(* IEC 61131-3 sources: daoli-st-library/DL_MathData (part 17) *)

(* ---- FC_DL_LinearScale.st ---- *)
(*==============================================================================
 * 组件名称 (Component)  : FC_DL_LinearScale
 * 所属子库 (Sublibrary) : DL_MathData
 * 当前版本 (Version)    : 1.0.0
 * 兼容性   (Platform)   : CODESYS 3.5 / TwinCAT 3 / 汇川 InoProShop / Machine Expert
 *                         仅依赖 Standard.library（ABS / MIN / MAX），全 REAL 运算
 * 功能描述 (Function)   : 模拟量原始码 → 工程量的线性标定。如 0..27648 对应 0..1.6MPa，
 *                         或 4..20mA 对应 0..100%。内置量程为零防御（除零保护）、
 *                         反向量程支持、输出双侧钳位、输入占量程百分比输出。
 *                         钳位判定使用浮点容差，不做浮点判等。
 * 开源溯源 (Origin)     : 原创实现。防御结构与模板库 05-algorithm-templates.md
 *                         的 FC_LinearScale 思路同源，按本库故障码体系重写并加严。
 * 依赖     (Depends)    : 无 DL_ 内部依赖
 * 说明     (Note)       : NaN / Inf 检测在纯 IEC 61131-3 中无标准手段（各平台对
 *                         比较运算返回值处理不一致），故 v1.0.0 不做该检测，
 *                         故障码 16#0001_0006 预留给支持 NaN 检测的平台版本。
 * 红线自检 (Redline)    : R1 ✓ 零全局变量表与外部变量引用 ｜ R2 ✓ 零物理 IO 地址直写
 *                         R3 ✓ 纯 IEC 61131-3 ｜ R4 ✓ 除零/排序/双侧钳位/容差判等（本轮 R4 样板）
 *                         R5 ✓ 全变量中英双语同行注释 ｜ R6 N/A（无状态机）｜ R7 N/A（无实例调用）
 * 修订历史 (Revision)   :
 *   2026-11-14  v1.0.0  首版入库（Phase 1 冷启动 · Level 0 批次）
 *============================================================================*)
FUNCTION FC_DL_LinearScale : REAL
VAR_INPUT
    fIn      : REAL;                 // 原始输入值 [raw] / Raw input value [raw]
    fInMin   : REAL := 0.0;          // 输入量程下限 [raw] / Input range low [raw]
    fInMax   : REAL := 27648.0;      // 输入量程上限 [raw] / Input range high [raw]
    fOutMin  : REAL := 0.0;          // 工程量下限 [EU] / Engineering range low [EU]
    fOutMax  : REAL := 100.0;        // 工程量上限 [EU] / Engineering range high [EU]
    bClamp   : BOOL := TRUE;         // 是否双侧钳位到工程量程 / Enable two-sided clamping
END_VAR
VAR_OUTPUT
    bValid   : BOOL;                 // 换算有效标志，FALSE 表示量程非法 / Conversion valid flag, FALSE means invalid range
    bClamped : BOOL;                 // 结果被钳位标志 / Result clamped flag
    fPercent : REAL;                 // 输入占量程百分比 [%]，可超 0..100 / Input as percent of span [%], may exceed 0..100
    uErrorId : UDINT;                // 故障码，0 = 无故障 / Error code, 0 = no error
END_VAR
VAR
    fSpanIn  : REAL;                 // 输入量程跨度 [raw]，可为负（反向标定） / Input span [raw], negative for reverse scaling
    fSpanOut : REAL;                 // 输出量程跨度 [EU]，可为负 / Output span [EU], may be negative
    fResult  : REAL;                 // 中间结果 [EU] / Intermediate result [EU]
    fNorm    : REAL;                 // 归一化比值 [0..1 附近]，无量纲 / Normalized ratio, dimensionless
    fOutLo   : REAL;                 // 输出下限，已排序 [EU] / Ordered output low limit [EU]
    fOutHi   : REAL;                 // 输出上限，已排序 [EU] / Ordered output high limit [EU]
    fBefore  : REAL;                 // 钳位前的结果快照，用于判定是否发生钳位 [EU] / Pre-clamp snapshot [EU]
END_VAR
VAR CONSTANT
    DL_FLOAT_EPS : REAL := 1.0E-6;   // 浮点判零容差 / Float zero tolerance
END_VAR

(*------------------------------------------------------------------------------
 * 段 1｜安全预置：任何异常路径下返回值落到工程量下限
 *      Safe preset: on every error path the return value falls back to the output low
 *-----------------------------------------------------------------------------*)
FC_DL_LinearScale := fOutMin;
bValid            := TRUE;
bClamped          := FALSE;
fPercent          := 0.0;
uErrorId          := 16#0000_0000;
fResult           := fOutMin;
fBefore           := fOutMin;

(*------------------------------------------------------------------------------
 * 段 2｜量程跨度计算 + 防除零（边界 B1 / B6）
 *      Span computation and divide-by-zero guard
 *      浮点判零用 ABS(..) <= EPS，禁止 fSpanIn = 0.0
 *      该段必须先于任何除法，fPercent 的计算建立在跨度已校验的前提上
 *-----------------------------------------------------------------------------*)
fSpanIn  := fInMax - fInMin;
fSpanOut := fOutMax - fOutMin;

IF ABS(fSpanIn) <= DL_FLOAT_EPS THEN
    bValid            := FALSE;
    uErrorId          := 16#0001_0002;
    FC_DL_LinearScale := fOutMin;
    RETURN;
END_IF

(*------------------------------------------------------------------------------
 * 段 3｜归一化与百分比（边界 B2）：反向量程天然支持
 *      Normalization and percentage: reverse ranges are supported by construction
 *      fInMax < fInMin 时 fSpanIn 为负，比值自动反向，0% 落在 fInMax 侧
 *-----------------------------------------------------------------------------*)
fNorm    := (fIn - fInMin) / fSpanIn;
fPercent := fNorm * 100.0;
fResult  := fOutMin + fNorm * fSpanOut;

(*------------------------------------------------------------------------------
 * 段 4｜输出边界排序（边界 B3）：钳位前必须先排序
 *      Output limit ordering before clamping
 *      若输出量程传反而不排序，钳位会把结果压到错误端点，现象是"钳位看似
 *      生效而输出全错"，这是本组件最隐蔽的失效模式
 *-----------------------------------------------------------------------------*)
fOutLo := MIN(fOutMin, fOutMax);
fOutHi := MAX(fOutMin, fOutMax);

(*------------------------------------------------------------------------------
 * 段 5｜双侧钳位（边界 B4/B5）：上下限成对出现，只用一侧是安全红线错误
 *      Two-sided clamping: both limits are mandatory, one-sided is a safety defect
 *      只做上限会让负向冲击直接打穿执行机构；钳位判定用容差而非不等号
 *-----------------------------------------------------------------------------*)
IF bClamp THEN
    fBefore := fResult;

    IF fResult < fOutLo THEN
        fResult := fOutLo;
    ELSIF fResult > fOutHi THEN
        fResult := fOutHi;
    END_IF

    IF ABS(fResult - fBefore) > DL_FLOAT_EPS THEN
        bClamped := TRUE;
    END_IF
END_IF

(*------------------------------------------------------------------------------
 * 段 6｜结果回写（边界 B7）：字面量均带小数点，全程 REAL，不混入 LREAL
 *      Result write-back: literals carry decimal points, REAL stays REAL
 *-----------------------------------------------------------------------------*)
FC_DL_LinearScale := fResult;
END_FUNCTION

(* ---- FC_DL_LineIntersection.st ---- *)
(*==============================================================================
 * 组件名称 (Component)  : FC_DL_LineIntersection
 * 所属子库 (Sublibrary) : DL_MathData
 * 当前版本 (Version)    : 1.0.0
 * 兼容性   (Platform)   : CODESYS 3.5 / TwinCAT 3 / 汇川 InoProShop / Machine Expert
 *                         仅依赖 Standard.library（ABS），全 LREAL 运算，无状态
 * 功能描述 (Function)   : 二维两直线（或两线段）交点求解。返回"是否存在唯一交点"的布尔量，
 *                         交点坐标与两个线段参数经状态输出给出，双通道并存的目的是让调用方
 *                         既能直接用作条件判断，也能拿到参数做端点命中判据。
 *                         用于视觉十字标定、皮带跑偏中心线求交、两台相机视场交叠区定位、
 *                         机器人平面两轴交汇点计算。
 *
 * 【失真与语义披露 / Distortion disclosure】
 *   1) 线段模式返回 FALSE 时 uErrorId = 0：业务上的"两段不相交"是正常判定结果，
 *      不是故障。若也置故障码，上位机会把正常判定当异常刷屏，真正的配置错误就被淹了。
 *   2) 重合直线归入平行类（16#0002_000D）：无穷多交点无法用单一坐标表达，
 *      与其随机给一个点，不如明确说"没有唯一交点"。线段模式下"平行且不共线"的两段
 *      永远不可能相交，属于正常业务判定，返回 FALSE 且不置码；只有重合（共线）才报码。
 *   3) 平行判据用绝对容差，而坐标量级到 1e6 时行列式 fDen 可到 1e12，因此 fEps 必须
 *      按坐标量级配置，经验式 fEps ≈ 1e-9 × 坐标量级²。用 1e-9 去判 1e12 量级的行列式，
 *      等于把平行判据关掉了。
 *   4) 本函数不检测 NaN/Inf：IEC 61131-3 无标准判据，强行判断会引入编译器方言。
 *
 * 开源溯源 (Origin)     : 原创实现（参考西门子 LGF 数学功能组中平面几何族的分类位置，
 *                         解析几何求交为公开数学方法，clean-room 独立实现）
 * 依赖     (Depends)    : 无 DL_ 内部依赖；Standard.library: ABS
 * 红线自检 (Redline)    : R1 ✓ 零全局变量表与外部变量引用 ｜ R2 ✓ 零物理 IO 地址直写
 *                         R3 ✓ 纯 IEC 61131-3（无指针、无厂商私有符号）
 *                         R4 ✓ 零长度线判据 + 容差规整 + 行列式判零 + 无交点显式清 0
 *                         R5 ✓ 全变量中英双语同行注释 ｜ R6 N/A（无状态机）｜ R7 N/A（无实例调用）
 * 修订历史 (Revision)   :
 *   2026-11-14  v1.0.0  首版入库（Phase 1 收口批次 · R3）
 *============================================================================*)
FUNCTION FC_DL_LineIntersection : BOOL
VAR_INPUT
    fX1         : LREAL;                  // 线 1 起点 X [mm] / Line 1 start X [mm]
    fY1         : LREAL;                  // 线 1 起点 Y [mm] / Line 1 start Y [mm]
    fX2         : LREAL;                  // 线 1 终点 X [mm] / Line 1 end X [mm]
    fY2         : LREAL;                  // 线 1 终点 Y [mm] / Line 1 end Y [mm]
    fX3         : LREAL;                  // 线 2 起点 X [mm] / Line 2 start X [mm]
    fY3         : LREAL;                  // 线 2 起点 Y [mm] / Line 2 start Y [mm]
    fX4         : LREAL;                  // 线 2 终点 X [mm] / Line 2 end X [mm]
    fY4         : LREAL;                  // 线 2 终点 Y [mm] / Line 2 end Y [mm]
    fEps        : LREAL := 1.0E-9;        // 平行判定容差（须按坐标量级配置）/ Parallel tolerance, scale with the coordinate range
    bSegmentMode: BOOL := FALSE;          // TRUE = 按线段求交，交点须落在两段内 / TRUE = segment mode
END_VAR
VAR_OUTPUT
    fX       : LREAL;                     // 交点 X [mm]，无交点时为 0 / Intersection X [mm], 0 when none
    fY       : LREAL;                     // 交点 Y [mm]，无交点时为 0 / Intersection Y [mm], 0 when none
    fT       : LREAL;                     // 线 1 参数 t，0 = 起点、1 = 终点 / Parameter along line 1
    fU       : LREAL;                     // 线 2 参数 u，0 = 起点、1 = 终点 / Parameter along line 2
    uErrorId : UDINT;                     // 故障码，0 = 无故障 / Error code, 0 = no error
END_VAR
VAR
    fDen  : LREAL;                        // 行列式分母 / Determinant denominator
    fDx1  : LREAL;                        // 线 1 方向 X 分量 [mm] / Line 1 direction X [mm]
    fDy1  : LREAL;                        // 线 1 方向 Y 分量 [mm] / Line 1 direction Y [mm]
    fDx2  : LREAL;                        // 线 2 方向 X 分量 [mm] / Line 2 direction X [mm]
    fDy2  : LREAL;                        // 线 2 方向 Y 分量 [mm] / Line 2 direction Y [mm]
    fEpsEff : LREAL;                      // 规整后的容差 / Normalised tolerance
    fTol  : LREAL;                        // 线段模式的参数区间容差 / Parameter tolerance in segment mode
    fNumT : LREAL;                        // t 的分子 / Numerator of t
    fNumU : LREAL;                        // u 的分子 / Numerator of u
    bLineDegenerate : BOOL;               // 任一线退化为点（起终点重合）/ Either line degenerated to a point
    bCoincident : BOOL;                   // 两线共线（重合），平行判定后的细分 / The two lines are coincident
END_VAR
VAR CONSTANT
    DL_LI_DEADBAND : LREAL := 1.0E-6;     // 零长度线判定容差 [mm] / Zero-length line tolerance [mm]
    DL_LI_EPS_MIN  : LREAL := 1.0E-12;    // 容差下限，防止把容差填成 0 / Tolerance floor
END_VAR

(*------------------------------------------------------------------------------
 * 段 1｜安全预置（边界 B6）：无交点时输出必须显式清 0，禁止依赖"局部变量默认值"
 *      Safe preset: outputs are explicitly zeroed, local defaults are never trusted
 *      部分平台的 FC 局部变量不保证每拍复位，靠默认值会让上一次的交点粘住
 *-----------------------------------------------------------------------------*)
FC_DL_LineIntersection := FALSE;
fX       := 0.0;
fY       := 0.0;
fT       := 0.0;
fU       := 0.0;
uErrorId := 16#0000_0000;

(*------------------------------------------------------------------------------
 * 段 2｜退化线检测（边界 B2）：起点终点重合/填反是最常见的标定配置错误，必须报码
 *      Degenerate-line check: start equal to end is the most common calibration mistake
 *      用曼哈顿距离判零长度：比平方和开方便宜，且对 LREAL 无溢出风险
 *-----------------------------------------------------------------------------*)
bLineDegenerate := ((ABS(fX2 - fX1) + ABS(fY2 - fY1)) <= DL_LI_DEADBAND)
                   OR ((ABS(fX4 - fX3) + ABS(fY4 - fY3)) <= DL_LI_DEADBAND);

IF bLineDegenerate THEN
    uErrorId := 16#0001_0001;
    RETURN;
END_IF

(*------------------------------------------------------------------------------
 * 段 3｜容差规整（边界 B1）：容差不能为 0 或负，否则平行判据失效
 *      Tolerance normalisation: zero or negative would disable the parallel test
 *-----------------------------------------------------------------------------*)
fEpsEff := fEps;

IF fEpsEff <= 0.0 THEN
    fEpsEff  := 1.0E-9;
    uErrorId := 16#0001_0001;
END_IF

IF fEpsEff < DL_LI_EPS_MIN THEN
    fEpsEff := DL_LI_EPS_MIN;
END_IF

(*------------------------------------------------------------------------------
 * 段 4｜方向向量与行列式（边界 B5）：分母只算一次，两条参数方程共用
 *      Direction vectors and determinant, computed once for both parametric equations
 *-----------------------------------------------------------------------------*)
fDx1 := fX2 - fX1;
fDy1 := fY2 - fY1;
fDx2 := fX4 - fX3;
fDy2 := fY4 - fY3;

fDen := (fDx1 * fDy2) - (fDy1 * fDx2);

(*------------------------------------------------------------------------------
 * 段 5｜平行/重合判定（边界 B3/B4）：无唯一交点
 *      Parallel or coincident: no unique intersection
 *      线段模式下"平行且不共线"的两段永远不相交，属正常业务判定，不置故障码；
 *      重合则有无穷多交点，仍是配置/数据问题，必须报码
 *      In segment mode, parallel non-collinear segments are a normal verdict, not a fault
 *-----------------------------------------------------------------------------*)
IF ABS(fDen) <= fEpsEff THEN

    bCoincident := (ABS(((fX3 - fX1) * fDy1) - ((fY3 - fY1) * fDx1)) <= fEpsEff);

    IF bSegmentMode AND (NOT bCoincident) THEN
        RETURN;
    END_IF

    uErrorId := 16#0002_000D;
    RETURN;

END_IF

(*------------------------------------------------------------------------------
 * 段 6｜参数求解：克拉默法则，分母在段 5 已判非零
 *      Parameter solution by Cramer's rule, the denominator was proven non-zero
 *-----------------------------------------------------------------------------*)
fNumT := (((fX3 - fX1) * fDy2) - ((fY3 - fY1) * fDx2));
fNumU := (((fX3 - fX1) * fDy1) - ((fY3 - fY1) * fDx1));

fT := fNumT / fDen;
fU := fNumU / fDen;

(*------------------------------------------------------------------------------
 * 段 7｜线段模式判定（边界 B3）：交点须落在两段的参数区间内
 *      Segment mode: the intersection must lie inside both parameter ranges
 *      端点命中算相交（容差取 fEpsEff 量级），否则相邻两段共端点时会被判成"不相交"；
 *      判定失败时 fT / fU 保留实际参数，便于上位机判断"差多远"，但坐标清 0
 *-----------------------------------------------------------------------------*)
IF bSegmentMode THEN

    fTol := fEpsEff;

    IF (fT < (0.0 - fTol)) OR (fT > (1.0 + fTol)) THEN
        (* 业务判定，不置故障码：线段不相交是正常结果 *)
        (* A business verdict, not a fault: disjoint segments are perfectly normal *)
        RETURN;
    END_IF

    IF (fU < (0.0 - fTol)) OR (fU > (1.0 + fTol)) THEN
        RETURN;
    END_IF

END_IF

(*------------------------------------------------------------------------------
 * 段 8｜交点求值（边界 B5）：一律由线 1 参数化，两式取平均会多引入一次误差
 *      Evaluate with line 1 only: averaging both equations adds error instead of removing it
 *-----------------------------------------------------------------------------*)
fX := fX1 + (fT * fDx1);
fY := fY1 + (fT * fDy1);

FC_DL_LineIntersection := TRUE;
END_FUNCTION

(* ---- FC_DL_LintToDintSat.st ---- *)
(*
    FC_DL_LintToDintSat —— LINT 到 DINT 双向域外饱和转换
    ------------------------------------------------------------------
    分类      : DL_MathData / Convert
    前缀      : FC_DL_
    版本      : 1.0.0
    溯源      : IEC 61131-3 标准语义的道莅防御性实现
                （接口语义由 IEC 61131-3 定义，内部委托平台内建 LINT_TO_DINT，
                  外围统一错误码 / 钳位 / 双语文档；clean-room 重写，
                  未复制任何闭源厂商源码，参考实现仅限 MIT/Apache 许可）
    平台      : 纯 IEC 61131-3，CODESYS / TwinCAT / InoProShop 通用
    作者      : 道莅代码库 · PLC编程专家（R17）
    ------------------------------------------------------------------
    功能说明  : 将 LINT 防御性转换为 DINT 并作为返回值输出，域内转换委托平台内建 LINT_TO_DINT；
                nIn 超 DINT 上界 2147483647 时饱和输出 2147483647 并置信息级 16#0001_0200；
                nIn 低于 DINT 下界 −2147483648 时饱和输出 −2147483648 并置信息级 16#0001_022D；
                下界输出采用计算式 -DL_DINT_MAX - 1，禁用负数字面量直写
                （部分编译器把负号解析为对一个越界正字面量取负，产生告警或错误结果）；
                极值比较采用双侧比较，禁用 ABS(nIn)（R55：有符号极值取绝对值会回绕漏判）；
                钳位方向：双侧饱和（−2147483648 ~ 2147483647），绝不回绕；
                纯整数域无 NaN/±INF 态，故无故障级路径（三个故障槽预留）。
    错误码    : 16#0001_0200 nIn 超 DINT 上界，已饱和至 2147483647——信息级，正常防御
                16#0001_022D nIn 低于 DINT 下界，已饱和至 −2147483648——信息级，正常防御
                16#0001_02EE 预留禁用（故障级，不得挪用）
                16#0001_02EF 预留禁用（故障级，不得挪用）
                16#0001_02F0 预留禁用（故障级，不得挪用）
    状态机    : R6 标注 N/A —— 本组件为纯函数无顺序状态机，无 CASE 可写，非法状态不可能出现，故以本节说明替代 ELSE 兜底
    修订记录  : 2026-11-16 v1.0.0 首次入库（R17）
*)
FUNCTION FC_DL_LintToDintSat : DINT
VAR_INPUT
    nIn : LINT; // 待转换 64 位有符号整数，建议域 ±9223372036854775807 [无量纲] / signed 64-bit integer to convert, suggested domain +/-9223372036854775807 [dimensionless]
END_VAR
VAR_OUTPUT
    eErr   : UDINT; // 错误码，0=正常 / error id, 0=ok
    bError : BOOL;  // 是否出错，eErr 非 0 时为 TRUE / error flag, TRUE when eErr is nonzero
    bValid : BOOL;  // 输出是否有效可用 / output valid flag
END_VAR
VAR CONSTANT
    DL_DINT_MAX_L : LINT := 2147483647;      // DINT 上界，用 LINT 承载以便域外比较 [无量纲] / DINT upper bound carried in LINT for out-of-domain comparison [dimensionless]
    DL_DINT_MIN_L : LINT := -2147483647 - 1; // DINT 下界，用 LINT 承载以便域外比较；下界值以计算式书写，避免负字面量解析歧义 [无量纲] / DINT lower bound carried in LINT, written as a computed expression to avoid negative literal parsing ambiguity [dimensionless]
    DL_DINT_MAX   : DINT := 2147483647;      // 上界饱和输出值 [无量纲] / upper saturation output [dimensionless]
    DL_DINT_ZERO  : DINT := 0;               // 返回值预置零（本件无故障路径） [无量纲] / preset zero, no fault path in this component [dimensionless]
END_VAR

// 段 1｜返回值与错误状态预置 / segment 1, preset return value and error status
FC_DL_LintToDintSat := DL_DINT_ZERO; // 预置 0（本件无故障级路径，仅作预置约定） [无量纲] / preset 0, no fault-level path in this component [dimensionless]
eErr   := 0;     // 预置无错误 / preset no error
bError := FALSE; // 预置无故障（本件无故障级路径） / preset no fault, no fault-level path here
bValid := FALSE; // 预置输出无效，通过双侧预判后置位 / preset invalid, set TRUE after both bound pre-checks

// 段 2｜上界预判与饱和 / segment 2, upper bound pre-check and saturation
IF nIn > DL_DINT_MAX_L THEN // 在 LINT 域先比较，超界值绝不送入内建转换 [无量纲] / compare in the LINT domain first, out-of-range values never reach the built-in conversion [dimensionless]
    FC_DL_LintToDintSat := DL_DINT_MAX; // 饱和输出 DINT 上界 2147483647 [无量纲] / saturate to the DINT upper bound 2147483647 [dimensionless]
    eErr := 16#0001_0200;               // 信息级：上溢饱和，正常防御 / info level: upper overflow saturated, normal defence
    bError := FALSE;                    // 信息级不置故障 / info level never raises fault
    bValid := TRUE;                     // 饱和值本身有效可用 / the saturated value itself is valid
    RETURN;                             // 饱和即出口，不调用内建转换 / saturation is the exit, built-in conversion not called
END_IF

// 段 3｜下界预判与饱和 / segment 3, lower bound pre-check and saturation
IF nIn < DL_DINT_MIN_L THEN // 双侧比较，禁用 ABS 单侧式（R55：有符号极值取绝对值会回绕） [无量纲] / two-sided comparison, single-sided ABS form forbidden, ABS of a signed extreme wraps around [dimensionless]
    FC_DL_LintToDintSat := -DL_DINT_MAX - 1; // 下界输出用计算式书写，等于 DINT 最小值 [无量纲] / lower bound output written as a computed expression, equal to the DINT minimum [dimensionless]
    eErr := 16#0001_022D;                    // 信息级：下溢饱和，正常防御 / info level: lower overflow saturated, normal defence
    bError := FALSE;                         // 信息级不置故障 / info level never raises fault
    bValid := TRUE;                          // 饱和值本身有效可用 / the saturated value itself is valid
    RETURN;                                  // 饱和即出口，不调用内建转换 / saturation is the exit, built-in conversion not called
END_IF

// 段 4｜域内委托转换（末段） / segment 4, in-domain delegated conversion (final)
FC_DL_LintToDintSat := LINT_TO_DINT(nIn); // 域内委托平台内建 LINT_TO_DINT，精确无损 [无量纲] / in-domain delegate to built-in LINT_TO_DINT, exact and lossless [dimensionless]
eErr   := 0;     // 域内无错误 / in-domain, no error
bError := FALSE; // 信息级不置故障 / info level never raises fault
bValid := TRUE;  // 域内输出有效可用 / in-domain output is valid
END_FUNCTION

(* ---- FC_DL_LintToLrealChk.st ---- *)
(*
    FC_DL_LintToLrealChk —— LINT 到 LREAL 精度告警防御转换
    ------------------------------------------------------------------
    分类      : DL_MathData / Convert
    前缀      : FC_DL_
    版本      : 1.0.0
    溯源      : IEC 61131-3 标准语义的道莅防御性实现
                （内部委托平台内建函数，外围统一错误码/钳位/双语文档；
                  未复制任何闭源厂商源码，参考实现仅限 MIT/Apache 许可）
    平台      : 纯 IEC 61131-3，CODESYS / TwinCAT / InoProShop 通用
    作者      : 道莅代码库 · PLC编程专家（R16）
    ------------------------------------------------------------------
    功能说明  : 将 LINT 输入防御性转换为 LREAL 并作为返回值输出；
                |nIn| 超过 2^53（9007199254740992，双精度浮点尾数 53 位精度极限）时，
                值照常转换输出，仅置信息级 16#0001_01CE 提示低位精度损失（bError=FALSE、bValid=TRUE）；
                钳位方向：无钳位（信息级仅记录，转换结果仍为最接近的可表值）；
                极值对称性防御：直接采用双侧比较 nIn > 上界 OR nIn < -下界，
                规避 ABS 对 LINT 最小值取绝对值的回绕未定义行为；
                域内转换委托平台内建 LINT_TO_LREAL 语义，不重实现数学内核；
                信息级码属正常防御：bError=FALSE、bValid=TRUE。
    错误码    : 16#0001_01CE |nIn| 超 2^53 精度极限，转换值低位可能失真——信息级，正常防御
                16#0001_01CF 预留禁用（信息级，不得挪用）
                16#0001_02A3 预留禁用（故障级，不得挪用）
                16#0001_02A4 预留禁用（故障级，不得挪用）
                16#0001_02A5 预留禁用（故障级，不得挪用）
    状态机    : R6 标注 N/A —— 本组件为纯函数无顺序状态机，无 CASE 可写，非法状态不可能出现，故以本节说明替代 ELSE 兜底
    修订记录  : 2026-11-16 v1.0.0 首次入库（R16）
*)
FUNCTION FC_DL_LintToLrealChk : LREAL
VAR_INPUT
    nIn : LINT; // 待转换输入 [无量纲] / input value to convert
END_VAR
VAR_OUTPUT
    eErr   : UDINT; // 错误码，0=正常 / error id, 0=ok
    bError : BOOL;  // 是否出错，eErr 非 0 时为 TRUE / error flag, TRUE when eErr is nonzero
    bValid : BOOL;  // 输出是否有效可用 / output valid flag
END_VAR
VAR CONSTANT
    DL_F53_MAX : LINT := 9007199254740992; // 双精度浮点尾数 53 位精度极限 2^53 [无量纲] / double-precision 53-bit mantissa precision limit 2^53
END_VAR

// 段 1｜返回值与错误状态预置 / segment 1, preset return value and error status
FC_DL_LintToLrealChk := 0.0; // 故障缺省返回 0 [无量纲] / fault default returns 0
eErr   := 0;     // 预置无错误 / preset no error
bError := FALSE; // 预置无故障（本组件无故障级路径） / preset no fault (no fault-level path in this component)
bValid := FALSE; // 预置无效，通过精度判定后置位 / preset invalid, set TRUE after precision check

// 段 2｜53 位精度极限判定与主体转换（末段） / segment 2, 53-bit precision limit check and main conversion (final)
IF (nIn > DL_F53_MAX) OR (nIn < -DL_F53_MAX) THEN
    FC_DL_LintToLrealChk := LINT_TO_LREAL(nIn); // 值照常转换（委托内建 _TO_ 语义） / convert as-is via built-in _TO_ conversion
    eErr := 16#0001_01CE; // 信息级：超 2^53 精度极限，低位可能失真，仅记录不钳位 / info level: beyond 2^53 precision limit, low bits may lose accuracy, record only
ELSE
    FC_DL_LintToLrealChk := LINT_TO_LREAL(nIn); // 域内委托平台内建 _TO_ 转换语义，精确无损 / in-domain delegate to built-in _TO_ conversion, exact lossless
    eErr := 0; // 域内无错误 / in-domain, no error
END_IF
bError := FALSE; // 信息级精度告警不置故障 / info-level precision notice never raises fault
bValid := TRUE;  // 域内或精度告警输出均有效可用 / in-domain or precision-noticed output is valid
END_FUNCTION

(* ---- FC_DL_LintToUdintSat.st ---- *)
(*
    FC_DL_LintToUdintSat —— LINT 到 UDINT 的双向饱和转换
    ------------------------------------------------------------------
    分类      : DL_MathData / Convert
    前缀      : FC_DL_
    版本      : 1.0.0
    溯源      : IEC 61131-3 类型定义的道莅防御性实现（LINT 64 位有符号 → UDINT 32 位无符号）；
                库内 FC_DL_LintToDintSat 只有「正向饱和」一个闸，本件补「负值落到无符号域」
                这一独立方向：两向的判据、出口与业务语义完全不同（负计数一律是组态错，
                超顶才是量程溢出）；双向闸、无损模式与错误分级 100% 自有；
                clean-room 重写，未复制任何闭源厂商源码，参考实现仅限 MIT/Apache 许可
    平台      : 纯 IEC 61131-3，CODESYS V3.5+ / TwinCAT 3 / InoProShop 通用
    作者      : 道莅代码库 · PLC编程专家（R19）
    ------------------------------------------------------------------
    功能说明  : 把 LINT 域内的计量/累计值安全落到 UDINT 域：负值饱和到 0，超顶饱和到
                4294967295；域内才委托内建 LINT_TO_UDINT（域外调用是三平台回绕行为
                不一致的根源，R56「无符号双分支钳位」同纪律）。
                核心防御：① 比较一律用 LINT 字面量常量，绝不把 UDINT 上限先当 UDINT 再比
                   （隐式升位在跨平台上有歧义）；
                ② 负向/正向各占一条信息码，方向可区分（R56 可 grep 化判据）；
                ③ bRequireLossless = TRUE 时任何饱和即判故障级 0327——计量与结算场景
                   不容许静默截断，宁可停机也不出错的数；
                ④ 域内路径零钳位、零额外比较开销。
                职责边界：有符号域内饱和（LINT→DINT）归 FC_DL_LintToDintSat，本件只管无符号落地。
    错误码    : 16#0001_0406 负向饱和（输入 < 0 → 0），组态错但已安全兜底——信息级，正常防御
                16#0001_0407 正向饱和（输入 > 4294967295 → 上限）——信息级，正常防御
                16#0001_0327 调用方要求无损（bRequireLossless = TRUE）却发生饱和——故障级，bValid = FALSE
                16#0001_0328 预留禁用（故障级，不得挪用）
                16#0001_0329 预留禁用（故障级，不得挪用）
    码位总账  : 16#0001_0406 用 / 16#0001_0407 用 ｜ 16#0001_0327 用 / 16#0001_0328 预留 / 16#0001_0329 预留
    状态机    : R6 标注 N/A —— 本组件为纯函数无顺序状态机，无 CASE 可写，非法状态不可能出现
    采样约定  : 本件无定时器、无沿检测、无状态；单拍纯计算，结论与任务周期无关。
    修订记录  : 2026-11-16 v1.0.0 首次入库（R19）
*)
FUNCTION FC_DL_LintToUdintSat : UDINT
VAR_INPUT
    liIn            : LINT := 0;              // 输入值 [无量纲]，全域 -2^63~2^63-1 / input value [dimensionless], full LINT domain
    bRequireLossless : BOOL := FALSE;         // TRUE = 发生任何饱和即判故障（计量/累计场景）/ TRUE turns any saturation into a fault for metering use
END_VAR
VAR_OUTPUT
    eErr            : UDINT;                  // 错误码，0=正常 / error id, 0=ok
    bError          : BOOL;                   // 故障标志，eErr 为故障级时 TRUE / error flag, TRUE on fault-level eErr
    bValid          : BOOL;                   // 返回值是否可用（饱和且要求无损时为 FALSE）/ return usable, FALSE when saturated in lossless mode
    bSatLow         : BOOL;                   // 负向饱和发生（输入 < 0）/ negative saturation occurred, input < 0
    bSatHigh        : BOOL;                   // 正向饱和发生（输入 > 4294967295）/ positive saturation occurred, input > 4294967295
END_VAR
VAR CONSTANT
    DL_UDINT_MAX_AS_LINT : LINT := 4294967295; // UDINT 上限的 LINT 形态 [无量纲] / the UDINT maximum expressed as LINT [dimensionless]
    DL_LINT_ZERO         : LINT := 0;          // 有符号零常量，避免裸字面量 [无量纲] / signed zero constant, avoids a bare literal [dimensionless]
    DL_UDINT_MAX         : UDINT := 16#FFFF_FFFF; // UDINT 上限值 [无量纲] / the UDINT maximum value [dimensionless]
    DL_UDINT_ZERO        : UDINT := 0;         // 无符号零常量 [无量纲] / unsigned zero constant [dimensionless]
END_VAR
VAR
    liWork          : LINT;                   // 输入副本，避免改动调用方数据 [无量纲] / input copy, never modifies caller data [dimensionless]
    uResult         : UDINT;                  // 转换结果中间量 [无量纲] / conversion result intermediate [dimensionless]
END_VAR

// 段 1｜返回值与错误状态预置 / segment 1, preset return value and error status
FC_DL_LintToUdintSat := DL_UDINT_ZERO;        // 故障缺省返回 0 / fault default returns zero
eErr := 0;                                    // 预置无错误 / preset no error
bError := FALSE;                              // 预置无故障 / preset no fault
bValid := FALSE;                              // 预置不可用，通过闸门后置位 / preset invalid, set TRUE after the gates
bSatLow := FALSE;                             // 预置未负向饱和 / preset no negative saturation
bSatHigh := FALSE;                            // 预置未正向饱和 / preset no positive saturation
uResult := DL_UDINT_ZERO;                     // 结果中间量清零 / clear the result intermediate

// 段 2｜负向闸门（负计数落到无符号域即组态错，先于正向判定）/ segment 2, negative gate
liWork := liIn;                               // 取入参副本参与比较 / copy the input for the comparisons
IF liWork < DL_LINT_ZERO THEN
    uResult := DL_UDINT_ZERO;                 // 负值饱和到 0 / saturate a negative value to zero
    bSatLow := TRUE;                          // 标记负向饱和 / flag the negative saturation
    eErr := 16#0001_0406;                     // 信息级：组态错但已安全兜底 / info level, configuration error handled safely
ELSE
    // 段 3｜正向闸门（用 LINT 字面量比较，绝不先转无符号再比）/ segment 3, positive gate
    IF liWork > DL_UDINT_MAX_AS_LINT THEN
        uResult := DL_UDINT_MAX;              // 超顶饱和到 4294967295 / saturate an overrun to the UDINT maximum
        bSatHigh := TRUE;                     // 标记正向饱和 / flag the positive saturation
        eErr := 16#0001_0407;                 // 信息级：量程溢出已兜底 / info level, range overrun handled safely
    ELSE
        // 段 4｜域内才委托内建（域外调用是三平台回绕不一致的根源）/ segment 4, delegate only inside the domain
        uResult := LINT_TO_UDINT(liWork);     // 域内无损转换 / lossless conversion inside the domain
        eErr := 0;                            // 域内无错误 / in-domain, no error
    END_IF
END_IF

// 段 5｜无损模式复核（要求无损却发生饱和即故障级）/ segment 5, lossless recheck
IF bRequireLossless AND (bSatLow OR bSatHigh) THEN
    eErr := 16#0001_0327;                     // 无损模式下发生饱和故障码 / saturation under lossless requirement
    bError := TRUE;                           // 置故障标志 / raise the error flag
    bValid := FALSE;                          // 返回值标记为不可用 / flag the return as unusable
    FC_DL_LintToUdintSat := uResult;          // 仍返回钳位值，便于 HMI 观察越界量 / still publish the clamped value so HMI can see the overrun
    RETURN;                                   // 出口 / exit
END_IF

// 段 6｜发布结果 / segment 6, publish the result
FC_DL_LintToUdintSat := uResult;              // 输出钳位后的无符号结果 [无量纲] / publish the clamped unsigned result [dimensionless]
bValid := TRUE;                               // 钳位或无损均可用 / usable either clamped or lossless
bError := FALSE;                              // 信息级不置故障 / info level never raises a fault
END_FUNCTION

(* ---- FC_DL_LnEx.st ---- *)
(*==============================================================================
 * 组件名称 (Component)  : FC_DL_LnEx
 * 所属子库 (Sublibrary) : DL_MathData
 * 当前版本 (Version)    : 1.0.0
 * 兼容性   (Platform)   : CODESYS 3.5 / TwinCAT 3 / 汇川 InoProShop / Machine Expert
 *                         仅依赖 Standard.library 的 LN 内建函数，
 *                         不重实现对数内核，无厂商数学方言依赖
 * 功能一句话 (Summary)  : 自然对数防御包装：fX <= 0 域闸门与非有限复检前置，
 *                         委托内建 LN，禁止 NaN / -Inf 穿透到下游联锁。
 * 功能描述 (Function)   : 对真数 fX 求自然对数。域闸门先行写死：
 *                         fX 非有限（NaN 用 x <> x 判据、无穷用 ABS(x) 超
 *                         有限性上界判据，均为库内既有写法）或 fX <= 0 时
 *                         不调内建、返回 0.0 并置码；fX = 0 在数学上趋于
 *                         -Inf，统一按域外拦截，不返回 -Inf；域内（fX > 0
 *                         且有限）委托内建 LN，结果再做一次非有限复检兜底。
 * 溯源     (Origin)     : IEC 61131-3 标准语义的道莅防御性实现
 *                         （接口语义由 IEC 61131-3 定义，clean-room 重写，
 *                         参考公开标准条款）
 * 码位     (Diag Codes) : 故障级 16#0001_0228（本件独占）：
 *                           fX <= 0 域外——LN(0) 数学上趋于 -Inf、LN(-x) 在
 *                           IEEE 754 下产生 NaN，本库统一拦截为「0.0 + 故障码」；
 *                         故障级 16#0001_0229（本件独占）：
 *                           输入或输出非有限（NaN / 无穷）拦截。
 * 类型裁定 (Type Note)  : 码位段 16#0001_xxxx 为全库共享 32 位段，WORD 容量不足，
 *                         故 eErr 采用 UDINT 承载（与库内 uErrorId : UDINT 惯例
 *                         一致，沿 R14 批 3 同一裁定）。
 * 依赖     (Depends)    : 无 DL_ 内部依赖；Standard.library: LN / ABS
 * 红线自检 (Redline)    : R1 ✓ 零全局变量与外部变量引用 ｜ R2 ✓ 零物理 IO 地址直写
 *                         R3 ✓ 纯 IEC 61131-3 ｜ R4 ✓ 域闸门先行 + 结果非有限复检
 *                         R5 ✓ 全变量中英双语同行注释
 *                         R6 N/A（纯函数，无 CASE/ENUM 状态机，按批 4 口径标 N/A）
 *                         R7 N/A（FC 为纯函数，无实例调用，头注释显式说明）
 * 防御行为声明 (Defense): ① fX <= 0 一律域外：LN(0) 极限为 -Inf，若放行会让
 *                           下游比较器拿到负无穷毒值，本库统一返回 0.0 +
 *                           故障码 16#0001_0228，与 IEEE/平台默认行为差异在此；
 *                         ② 非有限复检先行：NaN 判据 fX <> fX（NaN 与任何值
 *                           包括自身比较均为不等，库内既有写法）、无穷判据
 *                           ABS(fX) > 1.0E308，命中即不调内建、早退返回 0.0；
 *                         ③ 域内委托内建 LN 内核，结果非有限复检兜底
 *                           （防御纵深，正常域内不可能触发）；
 *                         ④ 两级闸门按「先非有限、后定义域」次序写死，
 *                           不可调换（NaN 参与任何大小比较均为 FALSE，
 *                           先判域会把 NaN 静默放行）；
 *                         ⑤ 1.0E308 有限性上界提为只读常量，禁魔法数；
 *                         ⑥ 浮点全程不用等号直比判数值相等，仅用 < > 与
 *                           NaN 自不等判据，符合浮点容差红线口径。
 * 修订历史 (Revision)   :
 *   2026-11-16  v1.0.0  首版入库（R14 批 4 · T0 快车道）
 *============================================================================*)
FUNCTION FC_DL_LnEx : LREAL
VAR_INPUT
    fX : LREAL; // 真数 [无量纲]，须 > 0 且有限 / Antilogarithm argument [dimensionless], must be > 0 and finite
END_VAR
VAR_OUTPUT
    eErr : UDINT; // 错误码，16#0001_0228=fX<=0 域外，16#0001_0229=非有限拦截，0=无事件 / Error code, 16#0001_0228=argument <= 0, 16#0001_0229=non-finite interception, 0=no event
END_VAR
VAR CONSTANT
    DL_LN_FINITE : LREAL := 1.0E308; // 有限性上界 [无量纲]，超界判无穷（库内既有写法）/ Finiteness bound, values beyond treated as infinity (library idiom)
END_VAR

(*------------------------------------------------------------------------------
 * 段 1｜返回值与错误码预置：先归零，任何早退路径都不会留下脏码
 *      Preset return value and error code so no early-exit path leaves a stale code
 *-----------------------------------------------------------------------------*)
FC_DL_LnEx := 0.0;   // 返回值预置 0.0（安全值，绝不输出 NaN / -Inf）/ Preset return to 0.0 (safe value, never NaN or -Inf)
eErr       := 16#0000_0000;   // 错误码预置无事件 / Preset error code to no event

(*------------------------------------------------------------------------------
 * 段 2｜非有限复检先行（防御声明②④）：次序写死——NaN 先于定义域，
 *      否则 NaN 会在大小比较中被静默放行
 *      Non-finite recheck first (defense notes 2 and 4): fixed order, NaN gate
 *      precedes the domain gate or NaN would silently pass the comparisons
 *-----------------------------------------------------------------------------*)
IF (fX <> fX) OR (ABS(fX) > DL_LN_FINITE) THEN
    eErr := 16#0001_0229;   // 故障码：输入非有限（NaN / 无穷），拦截早退 / Fault: non-finite input (NaN or infinity), intercepted
    RETURN;                 // 返回预置安全值 0.0 / Return preset safe value 0.0
END_IF

(*------------------------------------------------------------------------------
 * 段 3｜定义域闸门（防御声明①）：fX <= 0 域外（含 fX = 0 的 -Inf 趋近），
 *      返回 0.0 + 故障码，NaN / -Inf 绝不穿透到下游联锁
 *      Domain gate (defense note 1): fX <= 0 out of domain (including the -Inf
 *      limit at zero), returns 0.0 with fault code, no NaN or -Inf propagation
 *-----------------------------------------------------------------------------*)
IF fX <= 0.0 THEN
    eErr := 16#0001_0228;   // 故障码：真数 <= 0 域外，返回安全值 0.0 / Fault: argument <= 0 out of domain, safe value 0.0 returned
    RETURN;                 // 返回预置安全值 0.0，不产生 NaN / -Inf / Return preset safe value 0.0, no NaN or -Inf produced
END_IF

(*------------------------------------------------------------------------------
 * 段 4｜域内委托内建内核（防御声明③）：fX > 0 且有限，委托内建 LN
 *      In-domain delegation to the built-in kernel (defense note 3):
 *      fX > 0 and finite, delegate to the built-in LN
 *-----------------------------------------------------------------------------*)
FC_DL_LnEx := LN(fX);   // 委托内建 LN 内核，不自实现对数 / Delegate to the built-in LN kernel, no re-implementation

(*------------------------------------------------------------------------------
 * 段 5｜结果非有限复检（防御声明③）：域内正常不可能触发，兜底拦截
 *      Result finiteness recheck (defense note 3): unreachable in the normal
 *      domain, kept as a bottom-line interception
 *-----------------------------------------------------------------------------*)
IF (FC_DL_LnEx <> FC_DL_LnEx) OR (ABS(FC_DL_LnEx) > DL_LN_FINITE) THEN
    FC_DL_LnEx := 0.0;    // 兜底安全值 0.0 / Bottom-line safe value 0.0
    eErr := 16#0001_0229;   // 故障码：结果非有限拦截 / Fault: non-finite result intercepted
END_IF
END_FUNCTION

(* ---- FC_DL_Log10Safe.st ---- *)
// FC_DL_Log10Safe v1.0.0
// 开源溯源：来源 brOscatLib（EXP10 镜像件反演族） / URL https://github.com/iec-oscat-mirror / 许可证 MIT / 借鉴点 对数换算非正域饱和返回语义
(*==============================================================================
 * 功能描述: 安全 log10。输入 fX > 0 时返回 LN(fX)/LN(10)；fX <= 0 或非有限时
 *           返回 -3.402823e38 饱和值并置 bValid=FALSE（物理无效域安全侧）。
 * 接口契约: 输入 fX；输出 bValid 回执，返回值为 log10 结果。
 * 修订历史: 2026-11-23  v1.0.0  R74 首版
 *==============================================================================*)

FUNCTION FC_DL_Log10Safe : REAL
VAR_INPUT
    fX : REAL := 1.0;   // 对数自变量，域 > 0 [无量纲] / Logarithm argument, domain > 0
END_VAR
VAR_OUTPUT
    bValid : BOOL;      // 结果有效回执 [-] / Result validity receipt
END_VAR
VAR CONSTANT
    DL_L10_SAT : REAL := -3.402823E38;   // REAL 负向饱和哨兵值 [无量纲] / Negative saturation sentinel
    DL_L10_EPS : REAL := 1.0E-6;         // 判零容差 [无量纲] / Zero-test epsilon
END_VAR

(* —— 段 0：全路径赋值缺省（无效域安全侧） —— *)
bValid := FALSE;                            // 有效回执预清 / Validity preset
FC_DL_Log10Safe := DL_L10_SAT;              // 返回值缺省负饱和 / Result default negative saturation

(* —— 段 1：域闸与非有限闸（NaN 自反判 + 非正域拦截） —— *)
IF (fX <> fX) THEN                          // NaN 自反判（判等禁令唯一例外） / NaN self-reflexive test
    RETURN;                                 // 无效返回饱和 / Invalid, return saturation
END_IF
IF fX <= DL_L10_EPS THEN                    // 非正域（含判零容差）拦截 / Non-positive domain intercepted
    RETURN;                                 // 无效返回饱和 / Invalid, return saturation
END_IF
IF fX >= 3.0E38 THEN                        // 近 Inf 幅值闸 / Near-Inf gate
    RETURN;                                 // 无效返回饱和 / Invalid, return saturation
END_IF

(* —— 段 2：正常换算（LN(fX)/LN(10)，LN(10) 为常量无除零） —— *)
FC_DL_Log10Safe := LN(fX) / 2.302585093;    // log10 = LN(fX)/LN(10) / Logarithm base ten via natural log
bValid := TRUE;                             // 有效回执 / Validity receipt

END_FUNCTION

(* ---- FC_DL_LogBaseEx.st ---- *)
(*
    FC_DL_LogBaseEx —— 任意底数对数防御包装
    ------------------------------------------------------------------
    分类      : DL_MathData / Log
    前缀      : FC_DL_
    版本      : 1.0.0
    溯源      : IEC 61131-3 标准语义的道莅防御性实现
                （接口语义由 IEC 61131-3 定义，内部委托平台内建 LN，
                  外围统一错误码 / 钳位 / 双语文档；clean-room 重写，
                  未复制任何闭源厂商源码，参考实现仅限 MIT/Apache 许可）
    平台      : 纯 IEC 61131-3，CODESYS / TwinCAT / InoProShop 通用
    作者      : 道莅代码库 · PLC编程专家（R17）
    ------------------------------------------------------------------
    功能说明  : 返回以 fBase 为底的 fIn 对数，按换底公式 LN(fIn)/LN(fBase) 实现，
                两处对数均委托平台内建 LN，不重实现任何对数内核；
                非有限输入判为故障级 16#0001_02CD，返回 0.0 且 bValid=FALSE；
                定义域非法（fIn ≤ 0 或 fBase ≤ 0）判为故障级 16#0001_02CE，返回 0.0；
                底数退化（|fBase − 1| < 1.0E-6，含 fBase = 1）判为故障级 16#0001_02CF，
                返回 0.0（底数为 1 时对数无定义，贴近 1 时商发散，必须先拦不使用除法）；
                钳位方向：无钳位（三路故障均拦截并回缺省值）。
    错误码    : 16#0001_01EA 预留禁用（信息级，不得挪用）
                16#0001_01EB 预留禁用（信息级，不得挪用）
                16#0001_02CD 非有限输入（fIn 或 fBase 为 NaN / ±INF）——故障级，返回 0.0
                16#0001_02CE 定义域非法（fIn ≤ 0 或 fBase ≤ 0）——故障级，返回 0.0
                16#0001_02CF 底数退化（fBase = 1 或 |fBase − 1| < 1.0E-6）——故障级，返回 0.0
    状态机    : R6 标注 N/A —— 本组件为纯函数无顺序状态机，无 CASE 可写，非法状态不可能出现，故以本节说明替代 ELSE 兜底
    修订记录  : 2026-11-16 v1.0.0 首次入库（R17）
*)
FUNCTION FC_DL_LogBaseEx : REAL
VAR_INPUT
    fIn   : REAL; // 待求对数的真数（须 > 0） [无量纲] / logarithm argument (must be > 0) [dimensionless]
    fBase : REAL; // 对数底数（须 > 0 且 ≠ 1；=2.0 即 log2 用法） [无量纲] / logarithm base (must be > 0 and not 1; 2.0 yields log2) [dimensionless]
END_VAR
VAR_OUTPUT
    eErr   : UDINT; // 错误码，0=正常 / error id, 0=ok
    bError : BOOL;  // 是否出错，eErr 非 0 时为 TRUE / error flag, TRUE when eErr is nonzero
    bValid : BOOL;  // 输出是否有效可用 / output valid flag
END_VAR
VAR CONSTANT
    DL_LOG_FAULT_DEF  : REAL := 0.0;       // 故障缺省返回值 log10(1)=0 [无量纲] / fault default return value log10(1)=0 [dimensionless]
    DL_LOG_BASE_EPS   : REAL := 1.0E-6;    // 底数贴近 1 的判定容差（|fBase−1| < 该值视为退化） [无量纲] / base-near-1 tolerance, below means degenerate
    DL_FLOAT_EPS      : REAL := 1.0E-6;    // 浮点除子判定容差（除法前复判） [无量纲] / floating divisor tolerance, re-checked before division
    DL_REAL_INF_GUARD : LREAL := 4.0E38;   // REAL 域 ±INF 判定阈值，高于 REAL 最大有限值 3.402823E38 [无量纲] / REAL +/-INF guard above max finite REAL 3.402823E38
END_VAR
VAR
    fLnBase    : REAL; // 底数自然对数 LN(fBase) [无量纲] / natural logarithm of the base [dimensionless]
    bNonFinite : BOOL; // 非有限（NaN 或 ±INF）判定结果 / non-finite (NaN or +/-INF) detection result
END_VAR

// 段 1｜返回值与错误状态预置 / segment 1, preset return value and error status
FC_DL_LogBaseEx := DL_LOG_FAULT_DEF; // 故障缺省返回 0.0，对下游限幅链中性 [无量纲] / fault default 0.0, neutral for downstream limiting [dimensionless]
eErr   := 0;     // 预置无错误 / preset no error
bError := FALSE; // 预置无故障 / preset no fault
bValid := FALSE; // 预置输出无效，通过全部域门后置位 / preset invalid, set TRUE after all domain gates

// 段 2｜非有限防御闸 / segment 2, non-finite guard
bNonFinite := (fIn <> fIn) OR (fIn > DL_REAL_INF_GUARD) OR (fIn < -DL_REAL_INF_GUARD)
           OR (fBase <> fBase) OR (fBase > DL_REAL_INF_GUARD) OR (fBase < -DL_REAL_INF_GUARD); // 真数与底数双向非有限判定（NaN 自不等 + 安全幅值判 ±INF） [无量纲] / non-finite check on both argument and base (NaN by self-inequality, +/-INF by safe magnitude) [dimensionless]
IF bNonFinite THEN
    eErr := 16#0001_02CD; // 非有限输入故障码 / non-finite input fault id
    bError := TRUE;       // 置故障标志 / raise error flag
    bValid := FALSE;      // 输出不可用 / output not usable
    RETURN;               // 故障级提前返回，保持缺省 0.0 / early return on fault, keep default 0.0
END_IF

// 段 3｜定义域（域门）判定 / segment 3, domain gate
IF (fIn <= 0.0) OR (fBase <= 0.0) THEN
    eErr := 16#0001_02CE; // 定义域非法故障码（真数 ≤ 0 或底数 ≤ 0） [无量纲] / domain fault id, argument or base <= 0 [dimensionless]
    bError := TRUE;       // 置故障标志 / raise error flag
    bValid := FALSE;      // 输出不可用 / output not usable
    RETURN;               // 故障级提前返回，保持缺省 0.0 / early return on fault, keep default 0.0
END_IF

// 段 4｜底数退化闸（防 LN 除零发散） / segment 4, base degeneracy gate (prevents LN divide blow-up)
IF ABS(fBase - 1.0) < DL_LOG_BASE_EPS THEN // 底数贴近 1 时 LN(fBase) → 0，商将发散，必须先拦 [无量纲] / base near 1 makes LN(base) approach 0 and the quotient blow up, must gate first [dimensionless]
    eErr := 16#0001_02CF; // 底数退化故障码（fBase = 1 或贴近 1） / degenerate base fault id, fBase = 1 or near 1
    bError := TRUE;       // 置故障标志 / raise error flag
    bValid := FALSE;      // 输出不可用 / output not usable
    RETURN;               // 故障级提前返回，保持缺省 0.0 / early return on fault, keep default 0.0
END_IF

// 段 5｜除子整备与主体除法（末段） / segment 5, divisor preparation and main division (final)
fLnBase := LN(fBase); // 底数自然对数，委托平台内建 LN [无量纲] / natural logarithm of the base via built-in LN [dimensionless]
IF ABS(fLnBase) <= DL_FLOAT_EPS THEN // 除子复判（域闸之外的除法前第二道保险） [无量纲] / divisor re-check, second guard before division [dimensionless]
    eErr := 16#0001_02CF; // 除子趋零仍归入底数退化故障码 / near-zero divisor still reported as degenerate base
    bError := TRUE;       // 置故障标志 / raise error flag
    bValid := FALSE;      // 输出不可用 / output not usable
    RETURN;               // 除法前拦截，绝不执行除法 / blocked before division, division never executed
END_IF
FC_DL_LogBaseEx := LN(fIn) / fLnBase; // 换底公式主体，真数对数同样委托内建 LN [无量纲] / change-of-base body, argument logarithm also delegated to built-in LN [dimensionless]
eErr   := 0;     // 域内无错误 / in-domain, no error
bError := FALSE; // 信息级不置故障 / info level never raises fault
bValid := TRUE;  // 域内输出有效可用 / in-domain output is valid
END_FUNCTION

(* ---- FC_DL_LogDomainNormalize.st ---- *)
(*
  Name        : FC_DL_LogDomainNormalize
  Category    : DL_MathData
  Version     : 1.0.0
  Purpose     : 对数域归一化：pH/浓度/浊度等跨量级测量按 log 域映射到 0~1 线性度输出，含定义域与底数守卫；/ Normalize a wide-dynamic-range measurement into 0..1 via a log-domain mapping, with domain and base guards
  溯源        : 借 t1-1-oscat·math 的分类/参数域组织，clean-room 实现
  Boundary    : ① 定义域闸：fVal/fMin <= 0、fMax <= fMin、fBase <= 0 → 返回 0.0 哨兵（非故障级）；
                ② 底数闸：|LN(fBase)| < eps（即 fBase = 1）→ 对数退化除零 → 返回哨兵；
                ③ 跨度闸：|LN 域跨度| < eps → 返回哨兵（不产生 Inf）；
                ④ 非有限输入（NaN/Inf）拒收返回哨兵；⑤ xClamp 决定越界饱和或线性外推。
*)
FUNCTION FC_DL_LogDomainNormalize : LREAL
VAR_INPUT
    fVal     : LREAL := 1.0;                 (* 原始测量值（pH/浓度/浊度），域 > 0 [工程单位] / Raw measurement, must be > 0 *)
    fMin     : LREAL := 0.001;               (* 归一化下界（映射到 0.0），域 > 0 [工程单位] / Lower bound mapped to 0.0 *)
    fMax     : LREAL := 100.0;               (* 归一化上界（映射到 1.0），域 > fMin [工程单位] / Upper bound mapped to 1.0 *)
    fBase    : LREAL := 10.0;                (* 对数底，域 > 0 且 <> 1（典型 10 或 2.718）[-] / Log base, > 0 and not 1 *)
    xClamp   : BOOL := TRUE;                 (* TRUE = 输出饱和到 0..1；FALSE = 允许越界外推 [-] / Clamp output to 0..1 *)
END_VAR
VAR
    fLnBase : LREAL;                         (* LN(底数) 缓存 [-] / Cached LN of base *)
    fLnMin  : LREAL;                         (* 下界的底数域对数值 [-] / Log-domain value of lower bound *)
    fLnMax  : LREAL;                         (* 上界的底数域对数值 [-] / Log-domain value of upper bound *)
    fSpan   : LREAL;                         (* 对数域跨度 = fLnMax - fLnMin [-] / Log-domain span *)
    fNorm   : LREAL;                         (* 未钳位归一值 [-] / Unclamped normalized value *)
END_VAR
VAR CONSTANT
    DL_LDN_EPS : LREAL := 1.0E-6;            (* 定义域/底数/跨度判零容差（REAL 量级）[-] / Domain epsilon *)
    DL_LDN_ONE : LREAL := 1.0;               (* 归一上限常量 [-] / Normalized upper bound *)
    DL_LDN_ZERO : LREAL := 0.0;              (* 归一/哨兵零点常量 [-] / Zero constant *)
END_VAR

(* —— 段 1：全路径预置哨兵（未命中合法分支即输出 0.0，无旧值残留） —— *)
FC_DL_LogDomainNormalize := DL_LDN_ZERO;      (* 哨兵 0.0：还原方向不饱和，交由调用侧组态闸判有效性 / Sentinel 0.0, validity judged by caller *)

(* —— 段 2：非有限输入拒收（NaN 自反、Inf 差判，禁用近似阈值） —— *)
IF (fVal <> fVal) OR (fMin <> fMin) OR (fMax <> fMax) OR (fBase <> fBase) THEN
    RETURN;                                   (* NaN 拒收 / NaN rejected *)
END_IF
IF ((fVal - fVal) <> (fVal - fVal)) OR ((fMin - fMin) <> (fMin - fMin))
   OR ((fMax - fMax) <> (fMax - fMax)) OR ((fBase - fBase) <> (fBase - fBase)) THEN
    RETURN;                                   (* Inf 拒收（x-x 非零即非有限） / Inf rejected *)
END_IF

(* —— 段 3：定义域闸（每个参与换算的引脚单独覆盖，R151） —— *)
IF (fVal <= DL_LDN_ZERO) OR (fMin <= DL_LDN_ZERO) OR (fBase <= DL_LDN_ZERO) THEN
    RETURN;                                   (* 对数域要求正数输入 / Log domain requires positive inputs *)
END_IF
IF (fMax - fMin) <= DL_LDN_EPS THEN
    RETURN;                                   (* 上界须严格大于下界（差比较用容差，禁 = ） / Upper must exceed lower, tolerance compare *)
END_IF

(* —— 段 4：底数与跨度闸（除零唯一出入口） —— *)
fLnBase := LN(fBase);                         (* 自然对数缓存，仅算一次 / Natural log cached once *)
IF ABS(fLnBase) < DL_LDN_EPS THEN
    RETURN;                                   (* 底数 = 1：LOG 退化为除零 / Base 1 degenerates to division by zero *)
END_IF
fLnMin := LN(fMin) / fLnBase;                 (* 下界折算到底数域（除子已过闸） / Lower bound in base domain *)
fLnMax := LN(fMax) / fLnBase;                 (* 上界折算到底数域 / Upper bound in base domain *)
fSpan := fLnMax - fLnMin;                     (* 对数域跨度 / Log-domain span *)
IF ABS(fSpan) < DL_LDN_EPS THEN
    RETURN;                                   (* 跨度退化：不产生 Inf / Degenerate span, no Inf *)
END_IF

(* —— 段 5：归一换算 + 可选饱和（饱和前先算实值，非先钳后算） —— *)
fNorm := (LN(fVal) / fLnBase - fLnMin) / fSpan;   (* 线性内插：0 → fMin，1 → fMax / Linear interpolation in log domain *)
IF xClamp THEN
    IF fNorm < DL_LDN_ZERO THEN
        fNorm := DL_LDN_ZERO;                 (* 下限饱和 0.0 / Lower saturation *)
    ELSIF fNorm > DL_LDN_ONE THEN
        fNorm := DL_LDN_ONE;                  (* 上限饱和 1.0 / Upper saturation *)
    END_IF
END_IF
FC_DL_LogDomainNormalize := fNorm;            (* 返回归一值 / Return normalized value *)
END_FUNCTION

(* ---- FC_DL_LogEx.st ---- *)
(*
    FC_DL_LogEx —— 底 10 常用对数防御包装
    ------------------------------------------------------------------
    分类      : DL_MathData / Log
    前缀      : FC_DL_
    版本      : 1.0.0
    溯源      : IEC 61131-3 标准语义的道莅防御性实现
                （接口语义由 IEC 61131-3 定义，内部委托平台内建 LOG，
                  外围统一错误码 / 钳位 / 双语文档；clean-room 重写，
                  未复制任何闭源厂商源码，参考实现仅限 MIT/Apache 许可）
    平台      : 纯 IEC 61131-3，CODESYS / TwinCAT / InoProShop 通用
    作者      : 道莅代码库 · PLC编程专家（R17）
    ------------------------------------------------------------------
    功能说明  : 返回输入值的底 10 常用对数（IEC LOG 语义），内部委托平台内建 LOG，
                不重实现任何对数内核；
                非有限输入（NaN 或 ±INF）判为故障级 16#0001_02CA，返回 0.0 且 bValid=FALSE；
                定义域非法（输入 ≤ 0）判为故障级 16#0001_02CB，返回 0.0 且 bValid=FALSE；
                钳位方向：无钳位（两路故障均拦截并回缺省值，不做域内改造）。
    错误码    : 16#0001_01E8 预留禁用（信息级，不得挪用）
                16#0001_01E9 预留禁用（信息级，不得挪用）
                16#0001_02CA 非有限输入（NaN 或 ±INF）——故障级，返回 0.0
                16#0001_02CB 定义域非法（输入 ≤ 0）——故障级，返回 0.0
                16#0001_02CC 预留禁用（故障级，不得挪用）
    状态机    : R6 标注 N/A —— 本组件为纯函数无顺序状态机，无 CASE 可写，非法状态不可能出现，故以本节说明替代 ELSE 兜底
    修订记录  : 2026-11-16 v1.0.0 首次入库（R17）
*)
FUNCTION FC_DL_LogEx : REAL
VAR_INPUT
    fIn : REAL; // 待求对数的输入值（须 > 0） [无量纲] / input value whose logarithm is taken (must be > 0) [dimensionless]
END_VAR
VAR_OUTPUT
    eErr   : UDINT; // 错误码，0=正常 / error id, 0=ok
    bError : BOOL;  // 是否出错，eErr 非 0 时为 TRUE / error flag, TRUE when eErr is nonzero
    bValid : BOOL;  // 输出是否有效可用 / output valid flag
END_VAR
VAR CONSTANT
    DL_LOG_FAULT_DEF : REAL := 0.0;                         // 故障缺省返回值 log10(1)=0 [无量纲] / fault default return value log10(1)=0 [dimensionless]
    DL_REAL_INF_GUARD : LREAL := 4.0E38;                     // REAL 域 ±INF 判定阈值，高于 REAL 最大有限值 3.402823E38 [无量纲] / REAL +/-INF guard above max finite REAL 3.402823E38
END_VAR
VAR
    bNonFinite : BOOL; // 非有限（NaN 或 ±INF）判定结果 / non-finite (NaN or +/-INF) detection result
END_VAR

// 段 1｜返回值与错误状态预置 / segment 1, preset return value and error status
FC_DL_LogEx := DL_LOG_FAULT_DEF; // 故障缺省返回 0.0，即 log10(1)，对下游限幅链中性 [无量纲] / fault default 0.0, i.e. log10(1), neutral for downstream limiting [dimensionless]
eErr   := 0;     // 预置无错误 / preset no error
bError := FALSE; // 预置无故障 / preset no fault
bValid := FALSE; // 预置输出无效，通过域门后置位 / preset invalid, set TRUE after domain gate

// 段 2｜非有限防御闸 / segment 2, non-finite guard
bNonFinite := (fIn <> fIn) OR (fIn > DL_REAL_INF_GUARD) OR (fIn < -DL_REAL_INF_GUARD); // 非有限判定（NaN 自不等 + 安全幅值判 ±INF） [无量纲] / non-finite check (NaN by self-inequality, +/-INF by safe magnitude) [dimensionless]
IF bNonFinite THEN
    eErr := 16#0001_02CA; // 非有限输入故障码 / non-finite input fault id
    bError := TRUE;       // 置故障标志 / raise error flag
    bValid := FALSE;      // 输出不可用 / output not usable
    RETURN;               // 故障级提前返回，保持缺省 0.0 / early return on fault, keep default 0.0
END_IF

// 段 3｜定义域（域门）判定 / segment 3, domain gate
IF fIn <= 0.0 THEN
    eErr := 16#0001_02CB; // 定义域非法故障码（输入 ≤ 0） [无量纲] / domain fault id, input <= 0 [dimensionless]
    bError := TRUE;       // 置故障标志 / raise error flag
    bValid := FALSE;      // 输出不可用 / output not usable
    RETURN;               // 故障级提前返回，保持缺省 0.0 / early return on fault, keep default 0.0
END_IF

// 段 4｜主体计算（末段） / segment 4, main calculation (final)
FC_DL_LogEx := LOG(fIn); // 域内直接委托平台内建 LOG（底 10），不复检结果 [无量纲] / delegate to built-in LOG (base 10) in-domain, no re-check [dimensionless]
eErr   := 0;     // 域内无错误 / in-domain, no error
bError := FALSE; // 信息级不置故障 / info level never raises fault
bValid := TRUE;  // 域内输出有效可用 / in-domain output is valid
END_FUNCTION

(* ---- FC_DL_LogSafe.st ---- *)
(*
    FC_DL_LogSafe —— 自然对数 Safe 族防御包装（零/负拦截 + 下界钳 1E-300 + 委托内建）
    ------------------------------------------------------------------
    分类      : DL_MathData / Math-Log
    前缀      : FC_DL_
    版本      : 1.0.0
    来源标签  : iec-std-wrapper（T0）
    溯源      : IEC 61131-3 标准语义的道莅防御性实现
                （内部委托平台内建 LN，外围钳位/错误码/双语文档；
                  未复制任何闭源厂商源码）
    平台      : 纯 IEC 61131-3，CODESYS / TwinCAT / InoProShop 通用
    分工声明  : 与存量 FC_DL_LnEx / FC_DL_LogBaseEx 分工——LnEx 为任意底对数
                码位族，LogBaseEx 为换底包装；本件只做自然对数的 Safe 族口径
                （x<=0 判错误返回安全下界不返回 NaN + 下界钳 1E-300）。
    作者      : 道莅代码库 · PLC 编程专家（R57）
    ------------------------------------------------------------------
    功能说明  : 求输入的自然对数。四段式防御（R45）：NaN 双判据拦截归零早退；
                x<=0 判错误，返回安全下界 LN(1E-300) 不返回 NaN；0<x<1E-300
                钳到下界 1E-300 并置 bClamped；域内委托内建 LN；结果复检兜底。
                1E-300 量级依据：LN(1E-300) ≈ -690.7755278982 可表，
                LN(0) 与负数对数在 IEC 平台行为未定义，必须上游拦截。
    错误码    : 0000 正常 / 16#0002_0001 入参非有限已归零 / 16#0002_0003 x<=0 已按安全下界返回 / 16#0002_0002 下界钳位发生
    修订记录  : 2026-11-21 v1.0.0 首次入库（R57 批 2 · 序号 8）
*)
FUNCTION FC_DL_LogSafe : LREAL
VAR_INPUT
    lrIn : LREAL; // 输入实数 [无量纲]，定义域 大于零 / input real value [dimensionless], domain above zero
END_VAR
VAR_OUTPUT
    eErr     : UDINT; // 错误码，0 = 正常 / error code, zero is ok
    bError   : BOOL;  // 出错标志，eErr 非 0 时为真 / error flag, true when eErr is nonzero
    bValid   : BOOL;  // 结果是否为真实值，拦截/钳位降级时为假 / the result is the true value, false when degraded
    bClamped : BOOL;  // 本次调用发生下界钳位 [-] / a floor clamp happened this call
END_VAR
VAR
    lrUse : LREAL; // 钳位后的实际计算入参 [无量纲] / the clamped value fed to the kernel [dimensionless]
END_VAR
VAR CONSTANT
    DL_LOG_FLOOR : LREAL := 1E-300; // 下界钳位值 [无量纲]，LN(1E-300) 约 -690.78 可表 / the floor clamp, its log is representable
END_VAR

// 段 1｜返回值与错误状态预置安全值（四段式第一段，R45）/ segment 1, preset the return and error states
FC_DL_LogSafe := 0.0; // 返回值预置安全值 0.0 / preset the return to the safe zero
eErr     := 16#0000_0000; // 错误码预置正常 / preset the code to ok
bError   := FALSE; // 错误标志预置假 / preset the error flag false
bValid   := TRUE; // 有效标志预置真 / preset the valid flag true
bClamped := FALSE; // 钳位标志预置假 / preset the clamp flag false

// 段 2｜非有限拦截（双判据）：命中不调内建直接早退 / segment 2, the non finite interception
IF (lrIn <> lrIn) OR ((lrIn - lrIn) <> (lrIn - lrIn)) THEN // NaN 或无穷 / NaN or infinity
    eErr   := 16#0002_0001; // 信息级：输入非有限已归零 / informational, a non finite input zeroed
    bError := TRUE; // 置错误标志 / raise the error flag
    bValid := FALSE; // 输出不可用 / the output void
    RETURN; // 返回预置安全值 0.0 / return the preset safe zero
END_IF

// 段 3｜定义域闸门：x<=0 错误返回安全下界不返回 NaN；0<x<下界钳到下界 / segment 3, the domain gate
IF lrIn <= 0.0 THEN // 零或负 / zero or negative
    lrUse    := DL_LOG_FLOOR; // 按下界执行（返回 LN(1E-300) 而非 NaN）/ run at the floor, LN returned instead of NaN
    eErr     := 16#0002_0003; // 错误级：零负入参按安全下界返回 / error grade, a nonpositive input returned at the safe floor
    bError   := TRUE; // 置错误标志 / raise the error flag
    bValid   := FALSE; // 输出不可用（仅降级参考）/ the output void, degraded reference only
    bClamped := TRUE; // 置钳位标志 / raise the clamp flag
ELSIF lrIn < DL_LOG_FLOOR THEN // 正值但低于下界 / positive but below the floor
    lrUse    := DL_LOG_FLOOR; // 钳到下界 / clamp to the floor
    eErr     := 16#0002_0002; // 信息级：下界钳位发生 / informational, a floor clamp happened
    bError   := TRUE; // 置错误标志 / raise the error flag
    bValid   := FALSE; // 钳位结果非真实值 / the clamped result is not the true value
    bClamped := TRUE; // 置钳位标志 / raise the clamp flag
ELSE // 域内直通 / inside the domain
    lrUse := lrIn; // 直通 / passthrough
END_IF

// 段 4｜委托内建 LN（禁重实现数学内核）/ segment 4, delegation to the built-in LN
FC_DL_LogSafe := LN(lrUse); // 委托内建内核，除域已证为正 / delegate to the built-in kernel, the argument proven positive

// 段 5｜结果复检兜底（防御纵深，正常路径不可达）/ segment 5, the result recheck as defense in depth
IF (FC_DL_LogSafe <> FC_DL_LogSafe) OR ((FC_DL_LogSafe - FC_DL_LogSafe) <> (FC_DL_LogSafe - FC_DL_LogSafe)) THEN // 结果非有限 / a non finite result
    FC_DL_LogSafe := 0.0; // 兜底安全值 / the bottom-line safe value
    IF eErr = 16#0000_0000 THEN // 首事件优先置码 / the first event keeps the code
        eErr   := 16#0002_0001; // 信息级：结果非有限已归零 / informational, a non finite result zeroed
        bError := TRUE; // 置错误标志 / raise the error flag
        bValid := FALSE; // 输出不可用 / the output void
    END_IF
END_IF
END_FUNCTION

(* ---- FC_DL_LrcChecksum.st ---- *)
(*==============================================================================
 * 组件名称 (Component)  : FC_DL_LrcChecksum
 * 所属子库 (Sublibrary) : DL_MathData
 * 当前版本 (Version)    : 1.0.0
 * 兼容性   (Platform)   : CODESYS 3.5 / TwinCAT 3 / 汇川 InoProShop / Machine Expert
 *                         仅依赖 Standard.library（ABS / 显式类型转换），无厂商方言
 * 功能描述 (Function)   : Modbus ASCII 模式的 LRC（纵向冗余校验）计算。
 *                         把地址、功能码、数据字节按无符号 8 位累加，
 *                         取二进制补码（256 - 累加和 的低 8 位）作为校验值。
 *                         用于电表、称重仪表、老式温控器等仍走 ASCII 模式
 *                         设备的收帧校验。
 *
 * 【帧边界声明 / Frame-boundary declaration（边界 B1）】
 *   **冒号 16#3A 与回车换行 16#0D/16#0A 不参与计算。**
 *   误把帧头帧尾算进累加和，是现场 LRC 对不上的第一原因。
 *   输入必须传"解码后"的字节：先用 FC_DL_HexStringToBytes 把 ASCII 字符
 *   解码为字节数组，再把该数组传入本函数——两步调用顺序不可颠倒。
 *   若误传 ASCII 字符码（'0' = 16#30 而非 16#00），结果必然错。
 *
 * 【与 CRC 的关系 / Relation to CRC（边界 B5）】
 *   LRC 与 CRC-16 不可互算、不可互验。ASCII 模式用 LRC，RTU 模式用 CRC，
 *   同一设备切换模式时校验字段同时变。配套函数见 FC_DL_Crc16Modbus。
 *
 * 【大小写与字节序 / Case and byte order（边界 B6）】
 *   返回值是数值字节。转 ASCII 十六进制字符（"FB" 还是 "fb"）由组帧方
 *   决定，本函数不输出字符串、不规定大小写。
 *
 * 【使用前提与配套组件 / Prerequisites and companion（边界 B2）】
 *   本函数是无状态纯函数：不保存上一次的报文、不持有任何跨周期数据，
 *   可在任意任务周期安全调用，也支持同一扫描周期内对多路设备依次调用。
 *   上游配套为十六进制解码函数（先解码、后校验，见上方两步调用顺序）；
 *   下游如需 RTU 模式校验请改用 CRC-16 族函数，二者不可互验。
 *   收帧链路中冒号与回车换行必须在解码阶段被剥离，若上游解码函数
 *   配置为不剥帧，本函数的累加和将整体偏移，校验恒失败——
 *   该故障模式下 uSumLow 每次都对不上同一个值，可作为判据。
 *
 * 【验收向量 / Acceptance vectors（已实算复核，含逐字节和值分解）】
 *   V1  01 03 00 00 00 01（标准读保持寄存器请求）
 *       和值分解：01+03+00+00+00+01 = 16#05 → LRC = 16#FB
 *   V2  01 03 02 12 34（标准响应，寄存器值 1234）
 *       和值分解：01+03+02+12+34 = 16#4C → LRC = 16#B4
 *   V3  空报文（nLength = 0）→ 和 16#00 → 256-0 取模 → LRC = 16#00
 *       （正确值，非错误）
 *   V4  FF FF → 和 16#1FE，低 8 位 16#FE → 256-FE = 02 → LRC = 16#02
 *   V5  单字节 00 → 和 16#00 → LRC = 16#00
 *
 * 【两步调用顺序 / Two-step call sequence（边界 B2）】
 *   现场收帧的固定次序，不可颠倒：
 *     第一步：收到 ASCII 报文（含冒号与回车换行）后，先用配套的十六进制
 *             解码函数把报文体解码为字节数组（帧字符被剥离，不进数组）
 *     第二步：把解码后的字节数组与本函数要求的长度传入本函数，
 *             返回值即 LRC，与报文尾随的校验字符比对
 *   误传原始 ASCII 字符（如 '0' 的字符码 16#30 而非数值 16#00）时，
 *   累加和整体偏移，校验必然失败——这是现场第二常见错误。
 * 开源溯源 (Origin)     : 依 Modbus 应用协议规范（Modbus over Serial Line，
 *                         ASCII 传输模式定义）独立实现。OSCAT Network 校验
 *                         函数族仅提供"按协议分族、独立成函数"的组织方式参考
 *                         （EPL-2.0），未复制任何源码。
 * 依赖     (Depends)    : 无 DL_ 内部依赖（配套解码见 FC_DL_HexStringToBytes）
 * 红线自检 (Redline)    : R1 ✓ 零全局变量表与外部变量引用 ｜ R2 ✓ 零物理 IO 地址直写
 *                         R3 ✓ 纯 IEC 61131-3（显式 BYTE_TO_UDINT / UDINT_TO_BYTE）
 *                         R4 ✓ 长度钳位 + 下标双检 + 空报文兜底 + 宽类型防溢出
 *                         R5 ✓ 全变量中英双语同行注释 ｜ R6 N/A（无状态机）｜ R7 N/A（无实例调用）
 *
 * 【与 CRC 族函数的分工表 / Division of labour with the CRC family】
 *   传输模式      | 校验算法 | 本库配套函数           | 典型设备
 *   ASCII 串口    | LRC      | FC_DL_LrcChecksum      | 老式电表、称重仪表
 *   RTU 串口      | CRC-16   | FC_DL_Crc16Modbus      | 变频器、温控器
 *   以太网帧      | CRC-32   | FC_DL_Crc32Ethernet    | 固件下发、文件校验
 *   三者校验字段互不可算、互不可验；同一设备切换模式时校验字段同时变。
 * 修订历史 (Revision)   :
 *   2026-11-14  v1.0.0  首版入库（Phase 1 收口批次 · R3）
 *============================================================================*)
FUNCTION FC_DL_LrcChecksum : BYTE
VAR_IN_OUT
    aabyData  : ARRAY[0..255] OF BYTE;    // 参与校验的解码后字节（不含帧头帧尾） / Decoded payload bytes, framing excluded
END_VAR
VAR_INPUT
    nLength   : INT;                      // 字节数，合法域 0..256，越界自动钳位 / Byte count, range 0..256, clamped
END_VAR
VAR_OUTPUT
    uSumLow   : BYTE;                     // 累加和低 8 位（诊断用，LRC = 其补码） / Low byte of the sum for diagnostics
    uErrorId  : UDINT;                    // 故障码，0 = 无故障，16#0001_0001 = 长度越界已钳位 / Error code, 0 = no error, 0001_0001 = length clamped
END_VAR
VAR
    uSum      : UDINT;                    // 累加器，宽类型防中间溢出（禁止字节自加回绕） / Wide accumulator to avoid byte wrap-around
    nLenWork  : INT;                      // 钳位后的本地长度副本，不回写输入引脚 / Local clamped copy of the length
    nI        : INT;                      // 字节循环索引，值域 0..255 / Byte loop index, range 0..255
    nSumLowInt: INT;                      // 累加和低 8 位的整数形式，供补码运算 / Integer form of the low byte for two's complement math
END_VAR
VAR CONSTANT
    DL_LRC_MOD     : INT   := 256;        // 模 256，补码运算的模 / Modulus for two's complement math
    DL_LRC_BUF_MAX : INT   := 256;        // 缓冲上限，必须与数组维度一致 / Buffer limit, must match the array dimension
    DL_LRC_MASK    : UDINT := 16#0000_00FF; // 取低 8 位掩码 / Low-byte mask
END_VAR

(*------------------------------------------------------------------------------
 * 段 1｜安全预置：返回值与累加器归零，故障码清零
 *      Safe preset: return value and accumulator cleared, error code reset
 *      空报文（长度 0）是合法输入：和为 0，补码后 LRC = 16#00，
 *      这是正确值而非错误，不得报故障（边界 B3）。
 *      返回值先落 16#00 再进入计算：异常路径下不会返回未定义值，
 *      且 16#00 在补码口径下本就是合法的校验值（对应和值回绕到 0），
 *      与 CRC 族"返回值不得用 0 判错"的约定不同，此差异为算法本质。
 *-----------------------------------------------------------------------------*)
FC_DL_LrcChecksum := 16#00;
uSum              := 16#0000_0000;
uSumLow           := 16#00;
uErrorId          := 16#0000_0000;
nLenWork          := nLength;

(*------------------------------------------------------------------------------
 * 段 2｜长度防御（边界 B4）：钳位而非拒绝，让诊断链拿到可比对的值
 *      Length defence: clamp instead of reject, transient code on clamp
 *      负值 → 0；大于 256 → 256；均置 16#0001_0001（瞬时码）。
 *      选择钳位而非直接退回：现场排错时长度参数偶发抖动（比如上游
 *      把帧字符计入又纠正），直接退回会让诊断链断在第一步，
 *      钳位至少能给出一个"截断口径"的校验值供比对。
 *-----------------------------------------------------------------------------*)
IF nLenWork < 0 THEN
    nLenWork := 0;
    uErrorId := 16#0001_0001;
ELSIF nLenWork > DL_LRC_BUF_MAX THEN
    nLenWork := DL_LRC_BUF_MAX;
    uErrorId := 16#0001_0001;
END_IF

(*------------------------------------------------------------------------------
 * 段 3｜累加（边界 B4）：用 UDINT 宽类型累加，禁止依赖 BYTE 自加回绕——
 *      Accumulation in a wide UDINT accumulator
 *      部分平台对 BYTE 溢出回绕行为未定义，跨平台不可依赖。
 *      量级核算：256 字节全 0xFF 时累加和达 65280（16#FF00），
 *      UDINT 容量余量超过六万倍，本函数不存在累加溢出的可能，
 *      无需对累加器做饱和保护。
 *-----------------------------------------------------------------------------*)
IF nLenWork > 0 THEN

    FOR nI := 0 TO (nLenWork - 1) DO

        (* 数组下标上下界双检（红线 R4）：nLenWork ≤ 256 已保证 nI ≤ 255 *)
        (* Array index double check: nLenWork ≤ 256 guarantees nI ≤ 255 *)
        IF nI < DL_LRC_BUF_MAX THEN
            uSum := uSum + BYTE_TO_UDINT(aabyData[nI]);
        END_IF

    END_FOR;

END_IF

(*------------------------------------------------------------------------------
 * 段 4｜补码与回写：LRC = (256 - 累加和低 8 位) MOD 256
 *      Two's complement and write-back: LRC = (256 - low byte) MOD 256
 *      累加和低 8 位同步输出供诊断（对帧时可直接比对和值）。
 *      补码口径说明：本式等价于"按位取反加一后截取低 8 位"，
 *      但避免了取负运算，只依赖取模，跨平台行为完全一致。
 *      和值低 8 位为 0 时（含空报文与整字节回绕两种情况），
 *      LRC 均为 16#00，与 V3/V5 向量一致。
 *-----------------------------------------------------------------------------*)
uSumLow    := UDINT_TO_BYTE(uSum AND DL_LRC_MASK);
nSumLowInt := BYTE_TO_INT(uSumLow);

(* 显式 INT_TO_BYTE，MOD 已保证结果落在 0..255，无越界 *)
(* Explicit INT_TO_BYTE, MOD already bounds the result to 0..255 *)
FC_DL_LrcChecksum := INT_TO_BYTE((DL_LRC_MOD - nSumLowInt) MOD DL_LRC_MOD);

(*------------------------------------------------------------------------------
 * 段 5｜现场对拍指引（诊断用，无逻辑）
 *      On-site cross-check guidance for diagnostics, no logic here
 *      ① 收帧失败时先比对 uSumLow：与上位机侧算出的和值低 8 位一致，
 *        说明报文体一致、分歧在校验算法；不一致说明收到的字节本身有错，
 *        先查串口链路再查校验。
 *      ② 和值对、校验值不对：检查双方补码口径（本块为 256 减和取模，
 *        不是按位取反加一以外的变体）。
 *      ③ 和值偶尔对偶尔不对：多为帧字符混入或长度参数抖动，
 *        回查上游解码步骤的长度来源是否把帧字符计入了。
 *
 * 段 6｜自检向量断言说明（供单元测试与现场对拍，向量已实算复核）
 *      Self-check vector assertion notes, recomputed and verified
 *      V1  01 03 00 00 00 01 → 和 16#05 → uSumLow = 16#05、LRC = 16#FB
 *      V2  01 03 02 12 34   → 和 16#4C → uSumLow = 16#4C、LRC = 16#B4
 *      V3  空报文（长度 0）  → 和 16#00 → uSumLow = 16#00、LRC = 16#00
 *      V4  FF FF            → 和 16#1FE → uSumLow = 16#FE、LRC = 16#02
 *      V5  单字节 00         → 和 16#00 → uSumLow = 16#00、LRC = 16#00
 *-----------------------------------------------------------------------------*)
END_FUNCTION

(* ---- FC_DL_LrealSecToTime.st ---- *)
(*
    FC_DL_LrealSecToTime —— LREAL 秒到 TIME 防御转换（三路防御）
    ------------------------------------------------------------------
    分类      : DL_MathData / TimeConv
    前缀      : FC_DL_
    版本      : 1.0.0
    溯源      : IEC 61131-3 标准语义的道莅防御性实现
                （接口语义由 IEC 61131-3 定义，内部委托平台内建 LREAL_TO_TIME，
                  外围统一错误码 / 钳位 / 双语文档；clean-room 重写，
                  未复制任何闭源厂商源码，参考实现仅限 MIT/Apache 许可）
    平台      : 纯 IEC 61131-3，CODESYS / TwinCAT / InoProShop 通用
    作者      : 道莅代码库 · PLC编程专家（R17）
    ------------------------------------------------------------------
    功能说明  : 将 LREAL 秒数防御性转换为 TIME 并作为返回值输出，域内委托平台内建 LREAL_TO_TIME；
                非有限输入（NaN 或 ±INF）判为故障级 16#0001_02E2，返回 T#0S 且 bValid=FALSE；
                负值（TIME 无负语义）钳为 T#0S 并置信息级 16#0001_01F8；
                溢出预判先行：先在 LREAL 域与 4294967.295 s（对应 4294967295 ms）比较，
                超限直接饱和输出 T#49D17H2M47S295MS 并置信息级 16#0001_01F9，
                严禁把超限值乘 1000 后送进 LREAL_TO_TIME（先算后判必溢出）；
                钳位方向：下界钳 0 s，上界饱和至 TIME 域上限。
    错误码    : 16#0001_01F8 负秒输入（TIME 无负语义），已钳 T#0S——信息级，正常防御
                16#0001_01F9 秒数超 TIME 域上限（4294967.295 s），已饱和——信息级，正常防御
                16#0001_02E2 非有限输入（NaN 或 ±INF）——故障级，返回 T#0S
                16#0001_02E3 预留禁用（故障级，不得挪用）
                16#0001_02E4 预留禁用（故障级，不得挪用）
    状态机    : R6 标注 N/A —— 本组件为纯函数无顺序状态机，无 CASE 可写，非法状态不可能出现，故以本节说明替代 ELSE 兜底
    修订记录  : 2026-11-16 v1.0.0 首次入库（R17）
*)
FUNCTION FC_DL_LrealSecToTime : TIME
VAR_INPUT
    fSec : LREAL; // 秒数，有效域 0.0 ~ 4294967.295 s（负值钳 0，超限饱和） [s] / seconds, valid domain 0.0 .. 4294967.295 s, negative clamps, overflow saturates [s]
END_VAR
VAR_OUTPUT
    eErr   : UDINT; // 错误码，0=正常 / error id, 0=ok
    bError : BOOL;  // 是否出错，eErr 非 0 时为 TRUE / error flag, TRUE when eErr is nonzero
    bValid : BOOL;  // 输出是否有效可用 / output valid flag
END_VAR
VAR CONSTANT
    DL_SEC_MAX        : LREAL := 4294967.295;                     // TIME 域上限对应秒数（4294967295 ms） [s] / seconds equal to the TIME upper bound, 4294967295 ms [s]
    DL_SEC_MIN        : LREAL := 0.0;                             // 秒域下界 [s] / seconds lower bound [s]
    DL_MS_PER_SEC     : LREAL := 1000.0;                          // 秒转毫秒乘子（编译期常量） [ms/s] / seconds-to-milliseconds multiplier [ms/s]
    DL_TIME_MAX       : TIME  := T#49D17H2M47S295MS;              // TIME 域上限 4294967295 ms [ms] / TIME upper bound, 4294967295 ms [ms]
    DL_TIME_ZERO      : TIME  := T#0S;                            // TIME 零值（负值钳位与故障缺省） [ms] / TIME zero value, negative clamp and fault default [ms]
    DL_LREAL_HUGE     : LREAL := 1.7976931348623157E308;          // LREAL 最大有限幅值，超过即判 ±INF [无量纲] / max finite LREAL magnitude, beyond means +/-INF [dimensionless]
END_VAR
VAR
    bNonFinite : BOOL; // 非有限（NaN 或 ±INF）判定结果 / non-finite (NaN or +/-INF) detection result
END_VAR

// 段 1｜返回值与错误状态预置 / segment 1, preset return value and error status
FC_DL_LrealSecToTime := DL_TIME_ZERO; // 故障缺省返回 T#0S [ms] / fault default T#0S [ms]
eErr   := 0;     // 预置无错误 / preset no error
bError := FALSE; // 预置无故障 / preset no fault
bValid := FALSE; // 预置输出无效，通过三路闸后置位 / preset invalid, set TRUE after the three gates

// 段 2｜非有限防御闸 / segment 2, non-finite guard
bNonFinite := (fSec <> fSec) OR (fSec > DL_LREAL_HUGE) OR (fSec < -DL_LREAL_HUGE); // 非有限判定（NaN 自不等 + 最大有限幅值判 ±INF） [s] / non-finite check (NaN by self-inequality, +/-INF by max finite magnitude) [s]
IF bNonFinite THEN
    eErr := 16#0001_02E2; // 非有限输入故障码 / non-finite input fault id
    bError := TRUE;       // 置故障标志 / raise error flag
    bValid := FALSE;      // 输出不可用 / output not usable
    RETURN;               // 故障级提前返回，保持缺省 T#0S / early return on fault, keep default T#0S
END_IF

// 段 3｜负值闸与上界预判饱和 / segment 3, negative gate and upper-bound pre-check saturation
IF fSec < DL_SEC_MIN THEN
    FC_DL_LrealSecToTime := DL_TIME_ZERO; // 负值钳为 T#0S（TIME 无负语义） [ms] / clamp the negative value to T#0S, TIME has no negative semantics [ms]
    eErr := 16#0001_01F8;                 // 信息级：负秒已钳零，正常防御 / info level: negative seconds clamped to zero
    bError := FALSE;                      // 信息级不置故障 / info level never raises fault
    bValid := TRUE;                       // 钳位值本身有效可用 / the clamped value itself is valid
    RETURN;                               // 钳位即出口，不进入换算 / clamping is the exit, no scaling
END_IF
IF fSec > DL_SEC_MAX THEN // 在 LREAL 域先比较，先算后判必溢出 [s] / compare in the LREAL domain first, scaling before comparing would overflow [s]
    FC_DL_LrealSecToTime := DL_TIME_MAX; // 饱和至 TIME 域上限 T#49D17H2M47S295MS [ms] / saturate to the TIME upper bound T#49D17H2M47S295MS [ms]
    eErr := 16#0001_01F9;                // 信息级：秒数超上限已饱和，正常防御 / info level: seconds exceeded the upper bound and saturated
    bError := FALSE;                     // 信息级不置故障 / info level never raises fault
    bValid := TRUE;                      // 饱和值本身有效可用 / the saturated value itself is valid
    RETURN;                              // 饱和即出口，不进入换算 / saturation is the exit, no scaling
END_IF

// 段 4｜域内换算委托转换（末段） / segment 4, in-domain scaling and delegated conversion (final)
FC_DL_LrealSecToTime := LREAL_TO_TIME(fSec * DL_MS_PER_SEC); // 域内先乘常量 1000.0 转毫秒，再委托内建 LREAL_TO_TIME [ms] / in-domain multiply by the constant 1000.0 then delegate to built-in LREAL_TO_TIME [ms]
eErr   := 0;     // 域内无错误 / in-domain, no error
bError := FALSE; // 信息级不置故障 / info level never raises fault
bValid := TRUE;  // 域内输出有效可用 / in-domain output is valid
END_FUNCTION

(* ---- FC_DL_LrealToDintSat.st ---- *)
(*
    FC_DL_LrealToDintSat —— LREAL 到 DINT 向零截断饱和防御转换
    ------------------------------------------------------------------
    分类      : DL_MathData / Convert
    前缀      : FC_DL_
    版本      : 1.0.0
    溯源      : IEC 61131-3 标准语义的道莅防御性实现
                （内部委托平台内建函数，外围统一错误码/钳位/双语文档；
                  未复制任何闭源厂商源码，参考实现仅限 MIT/Apache 许可）
    平台      : 纯 IEC 61131-3，CODESYS / TwinCAT / InoProShop 通用
    作者      : 道莅代码库 · PLC编程专家（R16）
    ------------------------------------------------------------------
    功能说明  : 将 LREAL 输入防御性转换为 DINT 并作为返回值输出；
                非有限输入（NaN 或 ±INF）判为故障级 16#0001_0291，返回 0 且 bValid=FALSE；
                取整取向声明：向零截断（TRUNC 语义）后钳位，钳位按符号直接取界值；
                溢出预判先行（规避「先算后判」红线）：先在 LREAL 域判定越界并钳位，
                再对界值委托 TRUNC 向零截断，从而杜绝 TRUNC 越界未定义行为；
                越界时置信息级 16#0001_01C2（bError=FALSE、bValid=TRUE），输出钳位后防御值。
    错误码    : 16#0001_0291 非有限输入（NaN 或 ±INF）——故障级，返回 0
                16#0001_01C2 输入超 DINT 域，已按符号饱和钳位——信息级，正常防御
                16#0001_01C3 预留禁用（信息级，不得挪用）
                16#0001_0292 预留禁用（故障级，不得挪用）
                16#0001_0293 预留禁用（故障级，不得挪用）
    状态机    : R6 标注 N/A —— 本组件为纯函数无顺序状态机，无 CASE 可写，非法状态不可能出现，故以本节说明替代 ELSE 兜底
    修订记录  : 2026-11-16 v1.0.0 首次入库（R16）
*)
FUNCTION FC_DL_LrealToDintSat : DINT
VAR_INPUT
    fIn : LREAL; // 待转换输入 [无量纲] / input value to convert
END_VAR
VAR_OUTPUT
    eErr   : UDINT; // 错误码，0=正常 / error id, 0=ok
    bError : BOOL;  // 是否出错，eErr 非 0 时为 TRUE / error flag, TRUE when eErr is nonzero
    bValid : BOOL;  // 输出是否有效可用 / output valid flag
END_VAR
VAR CONSTANT
    DL_DINT_MAX   : LREAL := 2147483647.0;           // DINT 域上界，LREAL 承载 [无量纲] / DINT upper bound carried in LREAL
    DL_DINT_MIN   : LREAL := -2147483648.0;          // DINT 域下界，LREAL 承载 [无量纲] / DINT lower bound carried in LREAL
    DL_LREAL_HUGE : LREAL := 1.7976931348623157E308; // LREAL 最大有限幅值，超过即判 ±INF [无量纲] / max finite LREAL magnitude, beyond means +/-INF
END_VAR
VAR
    bNonFinite : BOOL; // 非有限（NaN 或 ±INF）判定结果 / non-finite (NaN or +/-INF) detection result
END_VAR

// 段 1｜返回值与错误状态预置 / segment 1, preset return value and error status
FC_DL_LrealToDintSat := 0; // 故障缺省返回 0 [无量纲] / fault default returns 0
eErr   := 0;     // 预置无错误 / preset no error
bError := FALSE; // 预置无故障 / preset no fault
bValid := FALSE; // 预置无效，通过防御闸后置位 / preset invalid, set TRUE after guard passes

// 段 2｜非有限防御闸 / segment 2, non-finite guard
bNonFinite := (fIn <> fIn) OR (fIn > DL_LREAL_HUGE) OR (fIn < -DL_LREAL_HUGE); // NaN 自不等判定，±INF 用安全幅值比较 [无量纲] / NaN by self-inequality, +/-INF by safe magnitude compare
IF bNonFinite THEN
    FC_DL_LrealToDintSat := 0; // 故障级返回 0 [无量纲] / fault level returns 0
    eErr   := 16#0001_0291;    // 非有限输入故障码 / non-finite input fault id
    bError := TRUE;            // 置故障标志 / set fault flag
    bValid := FALSE;           // 输出无效 / output invalid
    RETURN;                    // 立即返回 / immediate return
END_IF

// 段 3｜域判定先行钳位与向零截断主体计算（末段） / segment 3, domain-first clamp then truncate-toward-zero main conversion (final)
IF fIn > DL_DINT_MAX THEN
    FC_DL_LrealToDintSat := DL_DINT_MAX; // 正向钳至 DINT 上界（界值整数部分精确可表） / clamp to DINT upper bound (integer part exactly representable)
    eErr := 16#0001_01C2;                // 信息级：超上界已钳位 / info level: above upper bound, clamped
ELSIF fIn < DL_DINT_MIN THEN
    FC_DL_LrealToDintSat := DL_DINT_MIN; // 负向钳至 DINT 下界（界值整数部分精确可表） / clamp to DINT lower bound (integer part exactly representable)
    eErr := 16#0001_01C2;                // 信息级：超下界已钳位 / info level: below lower bound, clamped
ELSE
    FC_DL_LrealToDintSat := TRUNC(fIn); // 域内委托平台内建 TRUNC 向零截断 / in-domain delegate to built-in TRUNC toward zero
    eErr := 0; // 域内无错误 / in-domain, no error
END_IF
bError := FALSE; // 信息级钳位不置故障，故障分支已提前返回 / info-level clamp never raises fault, fault branch has returned
bValid := TRUE;  // 域内或钳位输出均有效可用 / in-domain or clamped output is valid
END_FUNCTION
